			// Cannel Status
			FOR i := MIN_CHANNEL TO MAX_CHANNEL DO	
				IF Force[i] THEN
					Status[i]								:= STATUS_ON;				
				ELSIF Receive[9-i] AND Receive[17-i] THEN   
					Status[i]								:= STATUS_OVERCURRENT;	
				ELSIF Receive[9-i] THEN                     
					Status[i]								:= STATUS_ON;
				ELSIF Receive[17-i] THEN                    
					Status[i]								:= STATUS_TRIP;
				ELSE                                        
					Status[i]								:= STATUS_OFF;
				END_IF                                      
			END_FOR		                                    
		                                                    
			// set collective triped bit                    
			FuseTripped										:= FALSE;
			FOR i := MIN_CHANNEL TO MAX_CHANNEL DO          
				IF Status[i] = STATUS_TRIP THEN             
					FuseTripped								:= TRUE;
					EXIT;
				END_IF
			END_FOR
			
			// interpret extended protoccol
			IF 	SendData[10] 
				OR 	SendData[11] 
			THEN			
				FOR i := MIN_CHANNEL TO MAX_CHANNEL DO // Voltage
					Temp									:= SHL(Temp,1) OR TO_BYTE(Receive[16+i]);
				END_FOR		  
				Voltage										:= Temp/16.0 + 16;
				FOR j := MIN_CHANNEL TO MAX_CHANNEL DO // Current[1-8]
					FOR i := MIN_CHANNEL TO MAX_CHANNEL DO    // bit shifting
						Temp								:= SHL(Temp,1) OR TO_BYTE(Receive[24+((j-1)*8)+i]);
					END_FOR		  
					Current[j]								:= Temp/16.0;
				END_FOR
			END_IF          
				
			UpdateCycle 									:= UpdateCycle + 1; 
			State 											:= 0;
		END_IF	
	END_CASE
	
(*****************************************************************)

PROPERTY PUBLIC baseClock : INT // MIN: 70 MAX: 200
GET
BaseClock := _BaseClock;
END_GET
SET
_BaseClock := LIMIT(70, BaseClock, 200);
State := -1;
END_SET
END_PROPERTY

METHOD reset : BOOL //Resetting tripped channel / Return TRUE as lons as FuseTripped = TRUE
VAR_INPUT
END_VAR
_InternReset													:= FuseTripped;
reset															:= TRUE;
END_METHOD

END_FUNCTION_BLOCK

// ---- POUs/Zeug/FB_FuseControl_1.TcPOU
FUNCTION_BLOCK FB_FuseControl_1
VAR_INPUT
	bResetChannels:	BOOL;
END_VAR
VAR_OUTPUT
	fbError:		FB_Error;
END_VAR
VAR
	bInFuse		AT %I* : BOOL;
	bOutFuse	AT %Q* : BOOL;
	
	fbDelay				: TON;
	
	fbRS				: RS;
END_VAR

fbRS(SET := bResetChannels, RESET1 := FALSE);
IF NOT bInFuse THEN
	fbError.M_Set(1, '48V-Sicherung hat ausgelöst', 0, E_ErrorIDs.eFuseTripped, E_ErrorSrcs.eFuse);
	fbDelay(IN := FALSE);
END_IF

IF fbRS.Q1 THEN
	fbDelay(IN := TRUE, PT := T#700MS);
	IF bInFuse THEN
		bOutFuse := TRUE;
	END_IF
	IF fbDelay.Q THEN
		fbDelay(IN := FALSE);
		bOutFuse := FALSE;
		fbRS(SET := bResetChannels, RESET1 := TRUE);
	END_IF
END_IF

END_FUNCTION_BLOCK

// ---- POUs/Aktorik/FB_VI_Light.TcPOU
FUNCTION_BLOCK FB_VI_Light
VAR_INPUT
	bLightOn				: BOOL;		// general light on
END_VAR
VAR_OUTPUT
	bError					: BOOL;		// error 
END_VAR
VAR_OUTPUT CONSTANT
	nIlluminationMaxBrightness : UINT := 511; // Firmware 92.51: 4095, Firmware 92.8: 511
END_VAR
VAR
	eResetHW			: E_ResetHW := E_ResetHW.INIT;	// Initial hardware reset to all illuminations
	stDeviceState		: ST_DeviceState;				// Basic state of device
	stLight				: ST_Light;						// Beckhoff illumination VI-R/P/B

	bErrorInternal		: BOOL;							// Error internal
	
	//light settings
	bIRActive						: BOOL  := TRUE; //activate infrared light
	nIRBrightnessPercent			: REAL := 10;	 //brightness of infrared light 
	bBlueActive						: BOOL := TRUE;	 //activate blue light
	nBlueBrightnessPercent			: REAL := 10;	 //brightness of blue light 
	bGreenActive					: BOOL := TRUE;  //activate green light
	nGreenBrightnessPercent			: REAL := 10;	 //brightness of green light 
	bOrangeActive					: BOOL := TRUE;	 //activate orange light
	nOrangeBrightnessPercent		: Real := 10;	 //brightness of orange light 
	
	nMaxTemperature					: SINT := 50;
	nTemperature					: SINT;
END_VAR

//state machine
CASE eResetHW OF 
	E_ResetHW.INIT:
		stLight.bEnable := FALSE;
		stLight.bReset := TRUE;		
		eResetHW := E_ResetHW.RESET_HW;
		RETURN;	
	E_ResetHW.RESET_HW:
		stLight.bReset := FALSE;
		eResetHW := E_ResetHW.DONE;
		RETURN;
	E_ResetHW.DONE:
		stLight.bEnable := TRUE;
		bErrorInternal := FALSE;
		IF NOT stDeviceState.Ready THEN
			bErrorInternal := TRUE;
			RETURN;
		ELSIF stDeviceState.Error THEN
			bLightOn := FALSE;
			stLight.bEnable := FALSE;
			eResetHW := E_ResetHW.INIT;
		END_IF

END_CASE

//-----------------------------------------------------------------------------------------------------------------
//set brightness and duration values for illumination 
stLight.channel[1].bActive		:= bIRActive;
stLight.channel[1].nBrightness	:= REAL_TO_UINT( nIRBrightnessPercent		* nIlluminationMaxBrightness / 100); // IR 
stLight.channel[2].bActive		:= bBlueActive;
stLight.channel[2].nBrightness	:= REAL_TO_UINT(nBlueBrightnessPercent	* nIlluminationMaxBrightness / 100); // blue 
stLight.channel[3].bActive		:= bGreenActive;
stLight.channel[3].nBrightness	:= REAL_TO_UINT(nGreenBrightnessPercent	* nIlluminationMaxBrightness / 100); // green 
stLight.channel[4].bActive		:= bOrangeActive;
stLight.channel[4].nBrightness	:= REAL_TO_UINT(nOrangeBrightnessPercent	* nIlluminationMaxBrightness / 100); // orange 

nTemperature := stLight.nTemperature;
  
//-----------------------------------------------------------------------------------------------------------------
// Automatic triggering
IF bLightOn AND nTemperature <= nMaxTemperature  THEN
//	IF  (NOT stLight.bActive AND nTemperature <= nMaxTemperature -10) TODO: Überhitzungsschutz als Hystherese
	stLight.bActive := TRUE;
	//bLightOn := FALSE; //TODO testen 
	
	bErrorInternal := FALSE;
	IF NOT stLight.bLightOn THEN
		bErrorInternal := TRUE;
	END_IF
ELSE
	stLight.bActive := FALSE;
END_IF

bError := stDeviceState.Error OR bErrorInternal;

METHOD PUBLIC SetIRGB : BOOL
VAR_INPUT
	nIRChannel		:	UINT;
	nRedChannel		:	UINT;
	nGreenChannel	:	UINT;
	nBlueChannel	:	UINT;
	nBrightness		:	REAL; 
END_VAR
nIRBrightnessPercent := (UINT_TO_REAL(nIrChannel)/255.0)*(nBrightness);
IF nIRChannel > 0 THEN
	bIRActive := TRUE;  
END_IF

nBlueBrightnessPercent := (UINT_TO_REAL(nBlueChannel)/255.0)*(nBrightness);  
IF nBlueChannel > 0 THEN
	bBlueActive := TRUE;  
END_IF
 
nGreenBrightnessPercent := (UINT_TO_REAL(nGreenChannel)/255.0)*(nBrightness); 
IF nGreenChannel > 0 THEN
	bGreenActive := TRUE;  
END_IF
 
nOrangeBrightnessPercent := (UINT_TO_REAL(nRedChannel)/255.0)*(nBrightness); 
IF nRedChannel > 0 THEN
	bOrangeActive := TRUE;  
END_IF
END_METHOD

METHOD SetWhiteLight : BOOL
VAR_INPUT
	nBrightness		: UINT := 100; 
END_VAR
SetIRGB(255, 255, 255, 255, nBrightness);
END_METHOD

END_FUNCTION_BLOCK

// ---- POUs/FB_ErrorCollector.TcPOU
FUNCTION_BLOCK FB_ErrorCollector
VAR_INPUT
END_VAR
VAR_OUTPUT
END_VAR
VAR
	i: INT;
END_VAR

METHOD M_NewError : BOOL
VAR_INPUT
	eID:	E_ErrorIDs;
	eSrc:	E_ErrorSrcs;
	sMsg: 	STRING;
END_VAR
FOR i := 0 TO HMI.nNumberErrors - 1 DO
	IF HMI.aErrors[i].nType = eID AND HMI.aErrors[i].nSource = eSrc THEN
		RETURN;
	END_IF
END_FOR

HMI.aErrors[HMI.nNumberErrors].nType := eID;
HMI.aErrors[HMI.nNumberErrors].nSource := eSrc;
HMI.aErrors[HMI.nNumberErrors].sMsg := sMsg;
HMI.nNumberErrors := HMI.nNumberErrors + 1;
HMI.bErrorChange := TRUE;
END_METHOD

METHOD M_QuitError : BOOL
VAR_INPUT
	eID:	E_ErrorIDs;
	eSrc:	E_ErrorSrcs;
END_VAR
FOR i := 0 TO HMI.nNumberErrors - 1 DO
	IF HMI.aErrors[i].nType = eID AND HMI.aErrors[i].nSource = eSrc THEN
		MEMSET(ADR(HMI.aErrors[i]), 0, SIZEOF(HMI.aErrors[i]));
		IF NOT (i = MAX_ERRORS - 1) THEN
			MEMMOVE(ADR(HMI.aErrors[i]), ADR(HMI.aErrors[i + 1]), SIZEOF(HMI.aErrors[i]) * HMI.nNumberErrors - i - 1);
			MEMSET(ADR(HMI.aErrors[HMI.nNumberErrors - 1]), 0, SIZEOF(HMI.aErrors[HMI.nNumberErrors - 1]));
		END_IF
		HMI.nNumberErrors := HMI.nNumberErrors - 1;
		HMI.bErrorChange := TRUE;
		EXIT;
	END_IF
END_FOR
END_METHOD

END_FUNCTION_BLOCK

// ---- POUs/Aktorik/FB_AxisCtrl.TcPOU
FUNCTION_BLOCK FB_AxisCtrl
VAR_INPUT
	eCommandIn:			E_AxesCmd;
	fPos:				LREAL;
	fVelo:				LREAL;
	bJogFw:				BOOL;
	bJogBw:				BOOL;
	
	bReset:				BOOL := TRUE;
END_VAR             	
VAR_OUTPUT
	bBusy:				BOOL;
	fbError:			FB_Error;
	bInRefPos AT %I* :	BOOL;
END_VAR             	
VAR_IN_OUT          	
	stAxis:				AXIS_REF;
END_VAR
VAR	
	eCommandAct:		E_AxesCmd;
	
	fbTimeout:			TON := (PT := T#90S);

//Achsen steuern
	fbMoveAbsolute:		MC_MoveAbsolute;
	fbMoveRelative:		MC_MoveRelative;
	fbJog:				MC_Jog;
	fbStop:				MC_Halt;
	fbReset:			MC_Reset;	
	fbSetPos:			MC_SetPosition;
END_VAR

A_Cycle();

CASE eCommandAct OF
	E_AxesCmd_IDLE:
		IF eCommandIn <> E_AxesCmd_IDLE THEN //neuer Auftrag
			eCommandAct := eCommandIn; //neuen Command speichern
		END_IF
		
	E_AxesCmd_MOVE_ABS:
		fbMoveAbsolute(Axis := stAxis, Execute := TRUE, Position := fPos, Velocity := fVelo);
		IF NOT fbMoveAbsolute.Busy THEN
			IF fbMoveAbsolute.Error THEN
				fbError.M_Set(fbMoveAbsolute.ErrorID, 'Achsen Fehler!', eCommandAct, eID := E_ErrorIDs.eAbsMove, eSrc := E_ErrorSrcs.eAxisCtrlPtp);
				eCommandAct := E_AxesCmd_ERROR;
			ELSE
				eCommandAct := E_AxesCmd_FINISHED;
			END_IF
			fbMoveAbsolute(Axis := stAxis, Execute := FALSE);
		ELSIF eCommandIn <> eCommandAct THEN
			fbMoveAbsolute(Axis := stAxis, Execute := FALSE);
			eCommandAct := E_AxesCmd_STOP;
		END_IF
		
	E_AxesCmd_MOVE_REL:
		fbMoveRelative(Axis := stAxis, Execute := TRUE, Distance := fPos, Velocity := fVelo);
		IF NOT fbMoveRelative.Busy THEN
			IF fbMoveRelative.Error THEN
				fbError.M_Set(fbMoveRelative.ErrorID, 'Achsen Fehler!', eCommandAct, eID := E_ErrorIDs.eRelMove, eSrc := E_ErrorSrcs.eAxisCtrlPtp);
				eCommandAct := E_AxesCmd_ERROR;
			ELSE
				eCommandAct := E_AxesCmd_FINISHED;
			END_IF
			fbMoveRelative(Axis := stAxis, Execute := FALSE);
		ELSIF eCommandIn <> eCommandAct THEN
			fbMoveRelative(Axis := stAxis, Execute := FALSE);
			eCommandAct := E_AxesCmd_STOP;
		END_IF
		
	E_AxesCmd_JOG:
		fbJog(Axis := stAxis, JogForward := bJogFw, JogBackwards := bJogFw, Mode := MC_JOGMODE_CONTINOUS, Velocity := fVelo);
		IF eCommandIn <> eCommandAct THEN
			fbJog(Axis := stAxis, JogForward := FALSE, JogBackwards := FALSE);
			eCommandAct := E_AxesCmd_IDLE;
		ELSIF fbJog.Error THEN
			fbError.M_Set(fbJog.ErrorID, 'Achsen Fehler!', eCommandAct, eID := E_ErrorIDs.eJog, eSrc := E_ErrorSrcs.eAxisCtrlPtp);
			eCommandAct := E_AxesCmd_ERROR;
		END_IF
	
	E_AxesCmd_STOP:
		fbStop(Axis := stAxis, Execute := TRUE);
		IF NOT fbStop.Busy THEN
			IF fbStop.Error THEN
				fbError.M_Set(fbStop.ErrorID, 'Achsen Fehler!', eCommandAct, eID := E_ErrorIDs.eJog, eSrc := E_ErrorSrcs.eAxisCtrlPtp);
				eCommandAct := E_AxesCmd_ERROR;
			ELSE
				eCommandAct := E_AxesCmd_FINISHED;
			END_IF
			fbStop(Axis := stAxis, Execute := FALSE);
		END_IF
		
	E_AxesCmd_FINISHED:
		IF eCommandIn = E_AxesCmd_IDLE THEN
			eCommandAct := E_AxesCmd_IDLE;
		END_IF
		
	E_AxesCmd_RESET:
		fbReset(Axis := stAxis, Execute := TRUE);
		IF NOT fbReset.Busy THEN
			IF fbReset.Error THEN
				fbError.M_Set(fbReset.ErrorID, 'Fehler bei Reset!', eCommandAct, eID := E_ErrorIDs.eResetAxis, eSrc := E_ErrorSrcs.eAxisCtrlPtp);
				eCommandAct := E_AxesCmd_ERROR;
			ELSE
				fbError.M_Reset();
				eCommandAct := E_AxesCmd_IDLE;
			END_IF
			fbReset(Axis := stAxis, Execute := FALSE);
		END_IF
		
	E_AxesCmd_ERROR:
		;
	
END_CASE

ACTION A_Cycle:

IF bReset THEN
	stAxis.ReadStatus();
	IF eCommandAct = E_AxesCmd_ERROR OR stAxis.Status.Error THEN
		eCommandAct := E_AxesCmd_RESET;				
	END_IF			
	bReset := FALSE;
END_IF

bBusy := eCommandAct <> E_AxesCmd_IDLE
	 AND eCommandAct <> E_AxesCmd_ERROR
	 AND eCommandAct <> E_AxesCmd_FINISHED;
END_ACTION

END_FUNCTION_BLOCK

// ---- POUs/Aktorik/FB_SimpleNcControl.TcPOU
FUNCTION_BLOCK FB_SimpleNcControl IMPLEMENTS I_NC_Ctrl
VAR CONSTANT
	VELO:				LREAL := 50;
END_VAR
VAR
	bEnable:			BOOL := TRUE;
	bReset:				BOOL;
	eState:				E_NC_State;
	bBusy:				BOOL;
	fbError:			FB_Error;

	
	rAxisX:				REFERENCE TO AXIS_REF;
	rAxisY:				REFERENCE TO AXIS_REF;
	rAxisZ:				REFERENCE TO AXIS_REF;
	
	fbAxisCtrlX:		FB_AxisCtrl;
	fbAxisCtrlY:		FB_AxisCtrl;
	fbAxisCtrlZ:		FB_AxisCtrl;
	
		
	fTargetX:			LREAL;
	fTargetY:			LREAL;
	fTargetZ:			LREAL;
		
	nRunState:			USINT; //0: Fall wählen; 10: nach oben, dann zum Ziel; 20: über Ziel fahren, dann senkrecht herunter //ZIEL: Gefahrenbereich umfahren
END_VAR

CASE eState OF	
	E_NC_State_INIT:
		IF __ISVALIDREF(rAxisX) AND __ISVALIDREF(rAxisY) AND __ISVALIDREF(rAxisZ) THEN			
			eState := E_NC_State_IDLE;
		END_IF

	E_NC_State_IDLE:
		;		
				
	E_NC_State_RUN:
		IF bEnable THEN
			CASE nRunState OF
				0:
					IF rAxisZ.NcToPlc.SetPos < MIN_MOVE_HEIGHT_Z AND (ABS(fTargetX - rAxisX.NcToPlc.SetPos) > 2 OR ABS(fTargetY - rAxisY.NcToPlc.SetPos) > 2) THEN
						nRunState := 10; //erst vertikal Gefahrenbereich verlassen, dann zum Ziel fahren
					ELSIF fTargetZ < MIN_MOVE_HEIGHT_Z AND (ABS(fTargetX - rAxisX.NcToPlc.SetPos) > 2 OR ABS(fTargetY - rAxisY.NcToPlc.SetPos) > 2) THEN
						nRunState := 20;
					ELSE
						nRunState := 11;
					END_IF
				
				10: //nach oben, dann zum Ziel
					fbAxisCtrlZ(stAxis := rAxisZ, eCommandIn := E_AxesCmd_MOVE_ABS, fPos := MIN_MOVE_HEIGHT_Z, fVelo := VELO);
					IF NOT fbAxisCtrlZ.bBusy THEN
						IF fbAxisCtrlZ.fbError.bError THEN
							fbError.M_Set(fbAxisCtrlZ.fbError.nErrorID, CONCAT('Achse Z: ', fbAxisCtrlZ.fbError.sErrorMsg), eState, eID := E_ErrorIDs.eAxisError, eSrc := E_ErrorSrcs.eAxisZ);
							eState := E_NC_State_ERROR;
						ELSE
							fbAxisCtrlZ(stAxis := rAxisZ, eCommandIn := E_AxesCmd_IDLE);
							nRunState := 0;
						END_IF
					END_IF
					
				11:
					fbAxisCtrlX(stAxis := rAxisX, eCommandIn := E_AxesCmd_MOVE_ABS, fPos := fTargetX, fVelo := VELO);
					fbAxisCtrlY(stAxis := rAxisY, eCommandIn := E_AxesCmd_MOVE_ABS, fPos := fTargetY, fVelo := VELO);
					fbAxisCtrlZ(stAxis := rAxisZ, eCommandIn := E_AxesCmd_MOVE_ABS, fPos := fTargetZ, fVelo := VELO);
					IF NOT fbAxisCtrlX.bBusy AND NOT fbAxisCtrlY.bBusy AND NOT fbAxisCtrlZ.bBusy THEN
						IF fbAxisCtrlX.fbError.bError THEN
							fbError.M_Set(fbAxisCtrlX.fbError.nErrorID, CONCAT('Achse X: ', fbAxisCtrlX.fbError.sErrorMsg), eState, eID := E_ErrorIDs.eAxisError, eSrc := E_ErrorSrcs.eAxisX);
							eState := E_NC_State_ERROR;
						ELSIF fbAxisCtrlY.fbError.bError THEN
							fbError.M_Set(fbAxisCtrlY.fbError.nErrorID, CONCAT('Achse Y: ', fbAxisCtrlY.fbError.sErrorMsg), eState, eID := E_ErrorIDs.eAxisError, eSrc := E_ErrorSrcs.eAxisY);
							eState := E_NC_State_ERROR;
						ELSIF fbAxisCtrlZ.fbError.bError THEN
							fbError.M_Set(fbAxisCtrlZ.fbError.nErrorID, CONCAT('Achse Z: ', fbAxisCtrlZ.fbError.sErrorMsg), eState, eID := E_ErrorIDs.eAxisError, eSrc := E_ErrorSrcs.eAxisZ);
							eState := E_NC_State_ERROR;
						ELSE
							fbAxisCtrlX(stAxis := rAxisX, eCommandIn := E_AxesCmd_IDLE);
							fbAxisCtrlY(stAxis := rAxisY, eCommandIn := E_AxesCmd_IDLE);
							fbAxisCtrlZ(stAxis := rAxisZ, eCommandIn := E_AxesCmd_IDLE);
							bBusy := FALSE;
							nRunState := 0;
							eState := E_NC_State_IDLE;
						END_IF
					END_IF
					
					
				20: //über Ziel fahren, dann senkrecht herunter
					fbAxisCtrlX(stAxis := rAxisX, eCommandIn := E_AxesCmd_MOVE_ABS, fPos := fTargetX, fVelo := VELO);
					fbAxisCtrlY(stAxis := rAxisY, eCommandIn := E_AxesCmd_MOVE_ABS, fPos := fTargetY, fVelo := VELO);
					fbAxisCtrlZ(stAxis := rAxisZ, eCommandIn := E_AxesCmd_MOVE_ABS, fPos := MIN_MOVE_HEIGHT_Z, fVelo := VELO);
					IF NOT fbAxisCtrlX.bBusy AND NOT fbAxisCtrlY.bBusy AND NOT fbAxisCtrlZ.bBusy THEN
						IF fbAxisCtrlX.fbError.bError THEN
							fbError.M_Set(fbAxisCtrlX.fbError.nErrorID, CONCAT('Achse X: ', fbAxisCtrlX.fbError.sErrorMsg), eState, eID := E_ErrorIDs.eAxisError, eSrc := E_ErrorSrcs.eAxisX);
							eState := E_NC_State_ERROR;
						ELSIF fbAxisCtrlY.fbError.bError THEN
							fbError.M_Set(fbAxisCtrlY.fbError.nErrorID, CONCAT('Achse Y: ', fbAxisCtrlY.fbError.sErrorMsg), eState, eID := E_ErrorIDs.eAxisError, eSrc := E_ErrorSrcs.eAxisY);
							eState := E_NC_State_ERROR;
						ELSIF fbAxisCtrlZ.fbError.bError THEN
							fbError.M_Set(fbAxisCtrlZ.fbError.nErrorID, CONCAT('Achse Z: ', fbAxisCtrlZ.fbError.sErrorMsg), eState, eID := E_ErrorIDs.eAxisError, eSrc := E_ErrorSrcs.eAxisZ);
							eState := E_NC_State_ERROR;
						ELSE
							fbAxisCtrlX(stAxis := rAxisX, eCommandIn := E_AxesCmd_IDLE);
							fbAxisCtrlY(stAxis := rAxisY, eCommandIn := E_AxesCmd_IDLE);
							fbAxisCtrlZ(stAxis := rAxisZ, eCommandIn := E_AxesCmd_IDLE);
							nRunState := 21;
						END_IF
					END_IF
				21:
					fbAxisCtrlZ(stAxis := rAxisZ, eCommandIn := E_AxesCmd_MOVE_ABS, fPos := fTargetZ, fVelo := VELO);
					IF NOT fbAxisCtrlZ.bBusy THEN
						IF fbAxisCtrlZ.fbError.bError THEN
							fbError.M_Set(fbAxisCtrlZ.fbError.nErrorID, CONCAT('Achse Z: ', fbAxisCtrlZ.fbError.sErrorMsg), eState, eID := E_ErrorIDs.eAxisError, eSrc := E_ErrorSrcs.eAxisZ);
							eState := E_NC_State_ERROR;
						ELSE
							fbAxisCtrlZ(stAxis := rAxisZ, eCommandIn := E_AxesCmd_IDLE);
							bBusy := FALSE;
							nRunState := 0;
							eState := E_NC_State_IDLE;
						END_IF
					END_IF
					
			END_CASE			
		ELSE
			eState := E_NC_State_ABORT;
		END_IF
		
	E_NC_State_ABORT:
		fbAxisCtrlX(stAxis := rAxisX);
		fbAxisCtrlY(stAxis := rAxisY);
		fbAxisCtrlZ(stAxis := rAxisZ);
		IF NOT fbAxisCtrlX.bBusy AND NOT fbAxisCtrlY.bBusy AND NOT fbAxisCtrlZ.bBusy THEN
			IF fbAxisCtrlX.fbError.bError THEN
				fbError.M_Set(fbAxisCtrlX.fbError.nErrorID, CONCAT('Achse X: ', fbAxisCtrlX.fbError.sErrorMsg), eState, eID := E_ErrorIDs.eAxisError, eSrc := E_ErrorSrcs.eAxisX);
				eState := E_NC_State_ERROR;
			ELSIF fbAxisCtrlY.fbError.bError THEN
				fbError.M_Set(fbAxisCtrlY.fbError.nErrorID, CONCAT('Achse Y: ', fbAxisCtrlY.fbError.sErrorMsg), eState, eID := E_ErrorIDs.eAxisError, eSrc := E_ErrorSrcs.eAxisY);
				eState := E_NC_State_ERROR;
			ELSIF fbAxisCtrlZ.fbError.bError THEN
				fbError.M_Set(fbAxisCtrlZ.fbError.nErrorID, CONCAT('Achse Z: ', fbAxisCtrlZ.fbError.sErrorMsg), eState, eID := E_ErrorIDs.eAxisError, eSrc := E_ErrorSrcs.eAxisZ);
				eState := E_NC_State_ERROR;
			ELSE
				eState := E_NC_State_IDLE;
			END_IF
		END_IF
		
	E_NC_State_ERROR:
		;
END_CASE

IF bReset THEN
	bReset := FALSE;
	fbError.M_Reset();
	IF eState = E_NC_State_ERROR THEN
		fbAxisCtrlX(stAxis := rAxisX, bReset := TRUE);
		fbAxisCtrlY(stAxis := rAxisY, bReset := TRUE);
		fbAxisCtrlZ(stAxis := rAxisZ, bReset := TRUE);
		eState := E_NC_State_IDLE;
	END_IF
END_IF

bBusy := eState <> E_NC_State_IDLE
	 AND eState <> E_NC_State_ERROR;

METHOD M_AxesReady : BOOL
VAR_INPUT
END_VAR

IF __ISVALIDREF(rAxisX) AND __ISVALIDREF(rAxisY) AND __ISVALIDREF(rAxisZ) THEN		
	rAxisX.ReadStatus();
	rAxisY.ReadStatus();
	rAxisZ.ReadStatus();
	IF rAxisX.Status.Operational AND rAxisY.Status.Operational AND rAxisZ.Status.Operational THEN
		M_AxesReady := TRUE;
	END_IF
END_IF
END_METHOD

METHOD M_AxisRef
VAR_INPUT
	rX: REFERENCE TO AXIS_REF;
	rY: REFERENCE TO AXIS_REF;
	rZ: REFERENCE TO AXIS_REF;
END_VAR

rAxisX REF= rX;
rAxisY REF= rY;
rAxisZ REF= rZ;
END_METHOD

METHOD M_CancelJob
fbAxisCtrlX(stAxis := rAxisX, eCommandIn := E_AxesCmd_IDLE);
fbAxisCtrlY(stAxis := rAxisY, eCommandIn := E_AxesCmd_IDLE);
fbAxisCtrlZ(stAxis := rAxisZ, eCommandIn := E_AxesCmd_IDLE);
eState := E_NC_State_ABORT;
END_METHOD

METHOD M_Cyclic
THIS^();

//fbAxesEnable(bEnableAxes := bEnable OR eState <> E_NC_State_IDLE, fOverride := AXES_OVERRIDE, stX := rAxisX, stY := rAxisY, stZ := rAxisZ);
fbAxisCtrlX(stAxis := rAxisX);
fbAxisCtrlY(stAxis := rAxisY);
fbAxisCtrlZ(stAxis := rAxisZ);
END_METHOD

METHOD M_NewJob
VAR_INPUT
	fTargetPosX	: LREAL;
	fTargetPosY	: LREAL;
	fTargetPosZ	: LREAL;
END_VAR
IF M_AxesReady() THEN
	IF eState = E_NC_State_IDLE THEN
		fTargetX := fTargetPosX;
		fTargetY := fTargetPosY;
		fTargetZ := fTargetPosZ;
		eState := E_NC_State_RUN;
		nRunState := 0;
		fbError.M_Reset();
	ELSIF eState = E_NC_State_RUN AND (fTargetX <> fTargetPosX OR fTargetY <> fTargetPosY OR fTargetZ <> fTargetPosZ) THEN	
		M_CancelJob();
	END_IF
ELSE
	fbError.M_Set(1, 'Achsen sind nicht bereit!', eState, eID := E_ErrorIDs.eAxesNotReady, eSrc := E_ErrorSrcs.eAxisCtrlPtp);
END_IF
END_METHOD


PROPERTY P_Busy : BOOL
GET
P_Busy := bBusy;
END_GET
END_PROPERTY

PROPERTY P_Enable : BOOL
SET
bEnable := P_Enable;
END_SET
END_PROPERTY

PROPERTY P_ErrID : UDINT
GET
P_ErrID := fbError.nErrorID;
END_GET
END_PROPERTY

PROPERTY P_ErrMsg : STRING
GET
P_ErrMsg := fbError.sErrorMsg;
END_GET
END_PROPERTY

PROPERTY P_Error : BOOL
GET
P_Error := fbError.bError;
END_GET
END_PROPERTY


PROPERTY P_Reset : BOOL
SET
bReset := P_Reset;
END_SET
END_PROPERTY

END_FUNCTION_BLOCK

// ---- GlobalTextList.TcGTLO
TEXTLIST GlobalTextList
  414 = 'Black'
  70 = 'SetPos X: %.1f'
  700 = 'SetPos Y: %.1f'
  460 = 'SetPos Z: %.1f'
  917 = 'Enable'
  132 = 'Enable Axes'
  155 = 'Endlage X'
  393 = 'Endlage X nci'
  637 = 'Endlage Y'
  359 = 'Endlage Z'
  401 = 'EndX %.1f'
  500 = 'EndY %.1f'
  660 = 'Job ID %.1f'
  870 = 'Job ID %i'
  277 = 'New Stone'
  145 = 'Quit'
  978 = 'Set Job'
  392 = 'Set new Job'
  910 = 'StartX %.1f'
  563 = 'StartY %.1f'
  588 = 'Velo %.1f'
  542 = 'X: %.1f mm'
  609 = 'X: %f mm'
  520 = 'Y: %.1f mm'
  252 = 'Y: %f mm'
  737 = 'Z: %.1f mm'
  431 = 'Z: %f mm'
END_TEXTLIST

// ---- VISUs/VISU.TcVIS
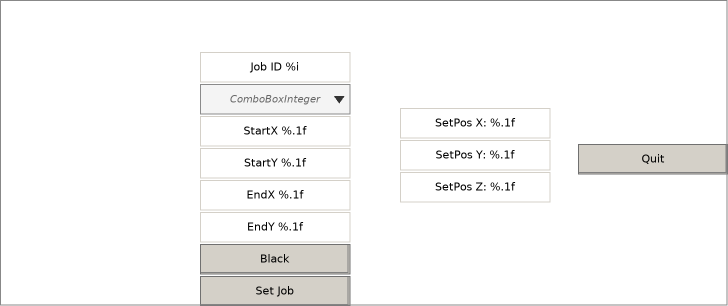
VISUALIZATION VISU  // 728x306
    Textfield (400,108 150x30), "SetPos X: %.1f", text variable: MAIN.fbIgorCtrl.fbPortal.aAxis[X].NcToPlc.SetPos
    Textfield (400,140 150x30), "SetPos Y: %.1f", text variable: MAIN.fbIgorCtrl.fbPortal.aAxis[Y].NcToPlc.SetPos
    Textfield (400,172 150x30), "SetPos Z: %.1f", text variable: MAIN.fbIgorCtrl.fbPortal.aAxis[Z].NcToPlc.SetPos
    Textfield (200,52 150x30), "Job ID %i", text variable: HMI.stJob.nJobID
        OnMouseClick: write HMI.stJob.nJobID via Default
    Textfield (200,180 150x30), "EndX %.1f", text variable: HMI.stJob.fDestPosX
        OnMouseClick: write HMI.stJob.fDestPosX via Default
    Textfield (200,116 150x30), "StartX %.1f", text variable: HMI.stJob.fStartPosX
        OnMouseClick: write HMI.stJob.fStartPosX via Default
    Textfield (200,148 150x30), "StartY %.1f", text variable: HMI.stJob.fStartPosY
        OnMouseClick: write HMI.stJob.fStartPosY via Default
    Textfield (200,212 150x30), "EndY %.1f", text variable: HMI.stJob.fDestPosY
        OnMouseClick: write HMI.stJob.fDestPosY via Default
    Button (200,276 150x30), "Set Job"
        tap HMI.bSetJob
    Button (578,144 150x30), "Quit"
        tap HMI.bQuit
    ComboBoxInteger (200,84 150x30), variable: HMI.stJob.eJobType
    Button (200,244 150x30), "Black"
        toggle HMI.stJob.bBlack
END_VISUALIZATION
